Fanuc KAREL source: kt00371.KL

-- PROVISIONAL review KL for V940-1; original PC SHA256 2b7e8b563051b6716ff98c5956129a184778bceedfe692d88df8908027e3dc53
-- Incomplete behavior may be omitted. Consult companion uncertainty JSON. Do not deploy.
PROGRAM KT00371
%NOLOCKGROUP
VAR
  R1 : REAL
  OUT : BOOLEAN
-- UNRESOLVED_DECL Y2 type=002018
BEGIN
  -- V9_ZERO_TABLE_METADATA_HINT layout=0001; no indexed target words; source/name/runtime held
  -- UNRESOLVED_PC offsets 5-16; opcodes 2E,23
  -- UNRESOLVED_PC offsets 21-35; opcodes 2E,22,9D,33,B2
  -- UNRESOLVED_PC offsets 40-63; opcodes 21,22,9D,33,B1,64,70,23
  -- UNRESOLVED_PC offsets 68-72; opcodes 7F
END KT00371
